Staubli VAL3: NewApp.dtx

public num nState
public num nAlarm
public string sAlarmMsg
public bool bStartCmd
public bool bStopCmd
public bool bPauseCmd
public bool bResetCmd
public bool bRunning
public num nCycleCount
public num nProdCount
